PROGRAM main
  VAR
    SCADA_LIGHTS_ON_CMD AT %QX0.0 : BOOL;
    SCADA_FAN_CMD AT %QX0.1 : BOOL;
    PUB_LIGHTS_MISMATCH AT %QX0.2 : BOOL;
    PUB_FAN_MISMATCH AT %QX0.3 : BOOL;
    PUB_LIGHTS_STATUS AT %QX0.4 : BOOL;
    PUB_FAN_STATUS AT %QX0.5 : BOOL;
    PUB_HEARTBEAT AT %QW0 : UINT;
    PUB_RECONNECT_COUNT AT %QW1 : UINT;
    LIGHTS_ON_CMD AT %QX100.0 : BOOL;
    FAN_CMD AT %QX100.1 : BOOL;
    LIGHTS_STATUS AT %IX100.0 : BOOL;
    FAN_STATUS AT %IX100.1 : BOOL;
    HEARTBEAT AT %IW100 : UINT;
    RECONNECT_COUNT AT %IW101 : UINT;
  END_VAR

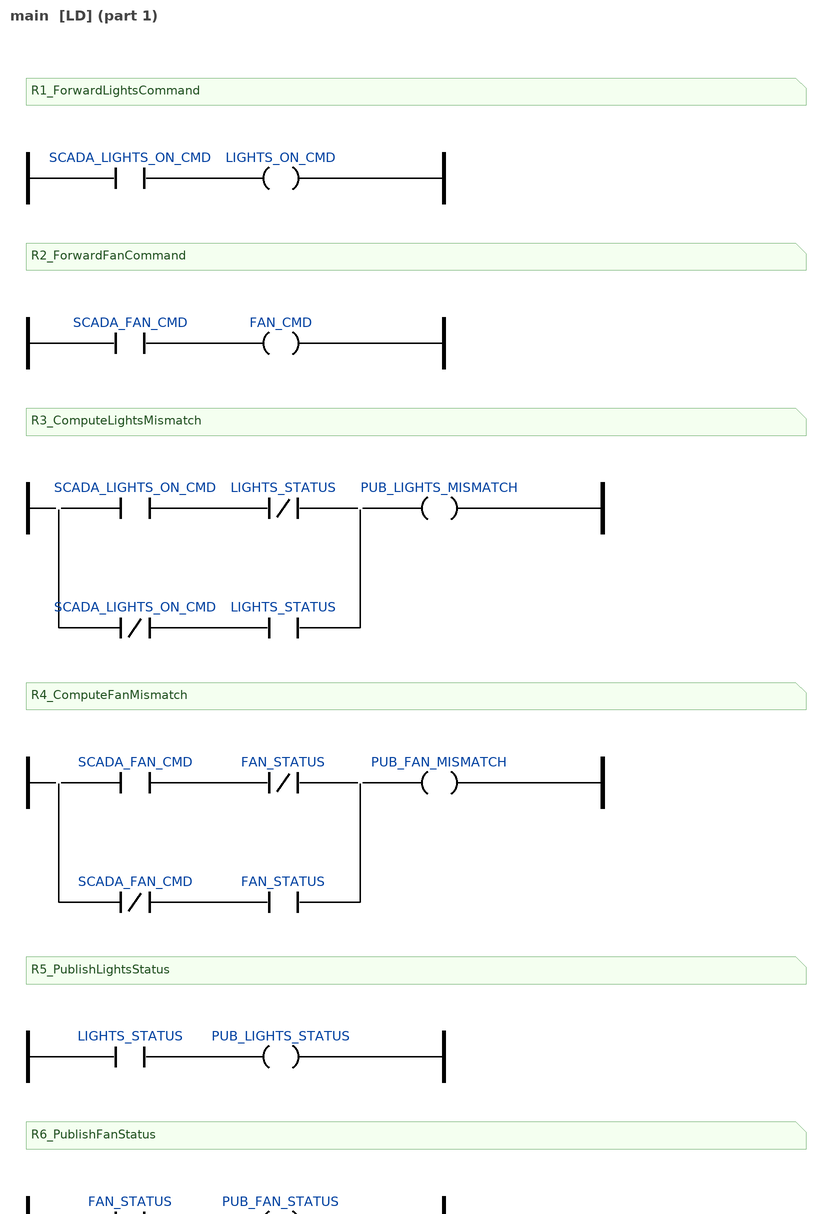
(* LD diagram, written out as Structured Text *)
(* R1_ForwardLightsCommand *)
LIGHTS_ON_CMD := SCADA_LIGHTS_ON_CMD;
(* R2_ForwardFanCommand *)
FAN_CMD := SCADA_FAN_CMD;
(* R3_ComputeLightsMismatch *)
PUB_LIGHTS_MISMATCH := NOT SCADA_LIGHTS_ON_CMD AND LIGHTS_STATUS OR SCADA_LIGHTS_ON_CMD AND NOT LIGHTS_STATUS;
(* R4_ComputeFanMismatch *)
PUB_FAN_MISMATCH := SCADA_FAN_CMD AND NOT FAN_STATUS OR NOT SCADA_FAN_CMD AND FAN_STATUS;
(* R5_PublishLightsStatus *)
PUB_LIGHTS_STATUS := LIGHTS_STATUS;
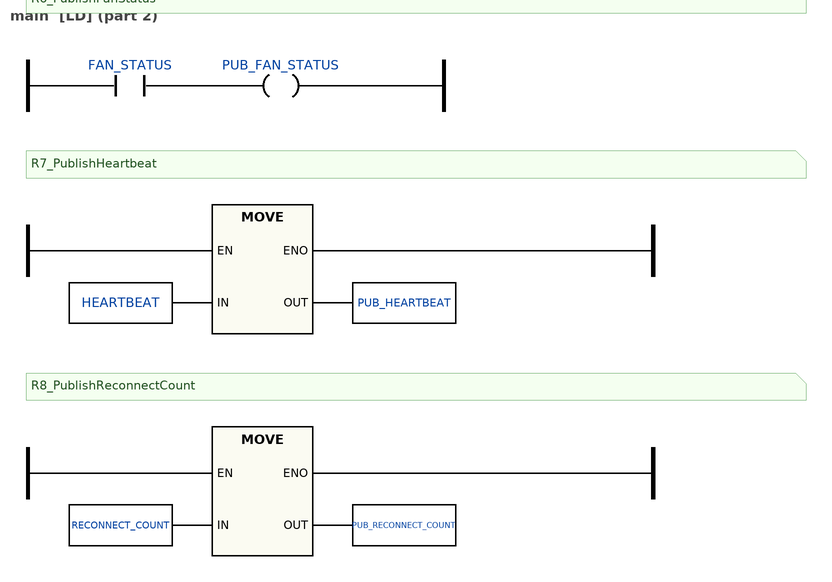
(* R6_PublishFanStatus *)
PUB_FAN_STATUS := FAN_STATUS;
(* R7_PublishHeartbeat *)
PUB_HEARTBEAT := HEARTBEAT;
(* R8_PublishReconnectCount *)
PUB_RECONNECT_COUNT := RECONNECT_COUNT;
END_PROGRAM
